FUNCTION_BLOCK PROCESS_IDENTIFICATION (* Offline identification prototype; see docs/adaptive/4diac-design.md *)
  (* Standard: 61499-2 *)
  (* Version 0.1, 2026-09-26, Guilherme *)
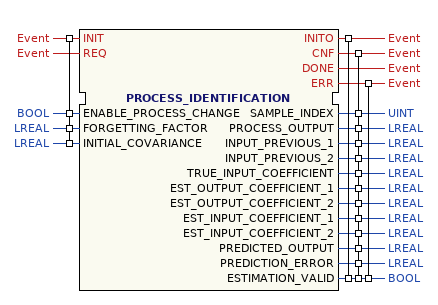
  EVENT_INPUT
    INIT WITH ENABLE_PROCESS_CHANGE, FORGETTING_FACTOR, INITIAL_COVARIANCE;
    REQ;
  END_EVENT
  EVENT_OUTPUT
    INITO WITH ESTIMATION_VALID;
    CNF WITH SAMPLE_INDEX, PROCESS_OUTPUT, INPUT_PREVIOUS_1, INPUT_PREVIOUS_2, TRUE_INPUT_COEFFICIENT, EST_OUTPUT_COEFFICIENT_1, EST_OUTPUT_COEFFICIENT_2, EST_INPUT_COEFFICIENT_1, EST_INPUT_COEFFICIENT_2, PREDICTED_OUTPUT, PREDICTION_ERROR, ESTIMATION_VALID;
    DONE;
    ERR WITH ESTIMATION_VALID;
  END_EVENT
  VAR_INPUT
    ENABLE_PROCESS_CHANGE : BOOL := FALSE;
    FORGETTING_FACTOR : LREAL := 1.0;
    INITIAL_COVARIANCE : LREAL := 10000.0;
  END_VAR
  VAR_OUTPUT
    SAMPLE_INDEX : UINT;
    PROCESS_OUTPUT : LREAL;
    INPUT_PREVIOUS_1 : LREAL;
    INPUT_PREVIOUS_2 : LREAL;
    TRUE_INPUT_COEFFICIENT : LREAL;
    EST_OUTPUT_COEFFICIENT_1 : LREAL;
    EST_OUTPUT_COEFFICIENT_2 : LREAL;
    EST_INPUT_COEFFICIENT_1 : LREAL;
    EST_INPUT_COEFFICIENT_2 : LREAL;
    PREDICTED_OUTPUT : LREAL;
    PREDICTION_ERROR : LREAL;
    ESTIMATION_VALID : BOOL;
  END_VAR
  FBS
    InputSequence : INPUT_SEQUENCE_REPLAY;
    OutputHistory : OUTPUT_HISTORY;
    SimulatedProcess : SECOND_ORDER_PROCESS;
    ParameterEstimator : RLS_PARAMETER_ESTIMATOR;
  END_FBS
  EVENT_CONNECTIONS
    INIT TO InputSequence.INIT;
    InputSequence.INITO TO OutputHistory.INIT;
    OutputHistory.INITO TO SimulatedProcess.INIT;
    SimulatedProcess.INITO TO ParameterEstimator.INIT;
    ParameterEstimator.INITO TO INITO;
    REQ TO InputSequence.REQ;
    InputSequence.CNF TO OutputHistory.REQ;
    OutputHistory.CNF TO SimulatedProcess.REQ;
    SimulatedProcess.CNF TO ParameterEstimator.REQ;
    ParameterEstimator.CNF TO OutputHistory.COMMIT;
    OutputHistory.ACK TO CNF;
    InputSequence.DONE TO DONE;
    ParameterEstimator.ERR TO ERR;
  END_CONNECTIONS
  DATA_CONNECTIONS
    ENABLE_PROCESS_CHANGE TO InputSequence.ENABLE_PROCESS_CHANGE;
    FORGETTING_FACTOR TO ParameterEstimator.FORGETTING_FACTOR;
    INITIAL_COVARIANCE TO ParameterEstimator.INITIAL_COVARIANCE;
    SimulatedProcess.PROCESS_OUTPUT TO ParameterEstimator.PROCESS_OUTPUT;
    SimulatedProcess.PROCESS_OUTPUT TO OutputHistory.CURRENT_OUTPUT;
    SimulatedProcess.PROCESS_OUTPUT TO PROCESS_OUTPUT;
    InputSequence.INPUT_PREVIOUS_1 TO SimulatedProcess.INPUT_PREVIOUS_1;
    InputSequence.INPUT_PREVIOUS_1 TO INPUT_PREVIOUS_1;
    InputSequence.INPUT_PREVIOUS_2 TO SimulatedProcess.INPUT_PREVIOUS_2;
    InputSequence.INPUT_PREVIOUS_2 TO INPUT_PREVIOUS_2;
    InputSequence.TRUE_INPUT_COEFFICIENT TO SimulatedProcess.TRUE_INPUT_COEFFICIENT;
    InputSequence.TRUE_INPUT_COEFFICIENT TO TRUE_INPUT_COEFFICIENT;
    InputSequence.SAMPLE_INDEX TO SAMPLE_INDEX;
    OutputHistory.OUTPUT_PREVIOUS_1 TO SimulatedProcess.OUTPUT_PREVIOUS_1;
    OutputHistory.OUTPUT_PREVIOUS_1 TO ParameterEstimator.OUTPUT_PREVIOUS_1;
    OutputHistory.OUTPUT_PREVIOUS_2 TO SimulatedProcess.OUTPUT_PREVIOUS_2;
    OutputHistory.OUTPUT_PREVIOUS_2 TO ParameterEstimator.OUTPUT_PREVIOUS_2;
    InputSequence.INPUT_PREVIOUS_1 TO ParameterEstimator.INPUT_PREVIOUS_1;
    InputSequence.INPUT_PREVIOUS_2 TO ParameterEstimator.INPUT_PREVIOUS_2;
    ParameterEstimator.EST_OUTPUT_COEFFICIENT_1 TO EST_OUTPUT_COEFFICIENT_1;
    ParameterEstimator.EST_OUTPUT_COEFFICIENT_2 TO EST_OUTPUT_COEFFICIENT_2;
    ParameterEstimator.EST_INPUT_COEFFICIENT_1 TO EST_INPUT_COEFFICIENT_1;
    ParameterEstimator.EST_INPUT_COEFFICIENT_2 TO EST_INPUT_COEFFICIENT_2;
    ParameterEstimator.PREDICTED_OUTPUT TO PREDICTED_OUTPUT;
    ParameterEstimator.PREDICTION_ERROR TO PREDICTION_ERROR;
    ParameterEstimator.ESTIMATION_VALID TO ESTIMATION_VALID;
  END_CONNECTIONS
END_FUNCTION_BLOCK
